(* IEC 61131-3 sources: rusty/tests/lit/single/arithmetic, 5 files *)

(* ---- addition.st ---- *)
// RUN: (%COMPILE %s && %RUN) | %CHECK %s
// CHECK: 10
FUNCTION main
    VAR
        x : DINT;
        y : DINT;
    END_VAR

    x := 5;
    y := 5;
    printf('%d$N', x + y);
END_FUNCTION

(* ---- integer_overflow.st ---- *)
// RUN: (%COMPILE %s && %RUN) | %CHECK %s
FUNCTION main
    VAR
        var_sint    : SINT;
        var_int     : INT;
        var_dint    : DINT;
        var_lint    : LINT;

        var_usint   : USINT;
        var_uint    : UINT;
        var_udint   : UDINT;
        var_ulint   : ULINT;
    END_VAR

    // Set max values
    // 8-bit [(2^7)-1]/[(2^8)-1]
    var_sint := 127;                    // Min: -128
    var_usint := 255;                   // Min: 0

    // 16-bit [(2^15)-1]/[(2^16)-1]
    var_int := 32767;                   // Min: -32768
    var_uint := 65535;                  // Min: 0

    // 32-bit [(2^31)-1]/[(2^31)-1]
    var_dint := 2147483647;             // Min: -2147483648
    var_udint := 4294967295;            // Min: 0

    // 64-bit [(2^63)-1]/[(2^64)-1]
    var_lint := 9223372036854775807;    // Min: -9223372036854775808
    var_ulint := 18446744073709551615;  // Min: 0

    // Print and check values
    printf('%d$N', var_sint);       // CHECK: 127
    printf('%d$N', var_int);        // CHECK-NEXT: 32767
    printf('%d$N', var_dint);       // CHECK-NEXT: 2147483647
    printf('%lld$N', var_lint);     // CHECK-NEXT: 9223372036854775807

    printf('%u$N', var_usint);      // CHECK-NEXT: 255
    printf('%u$N', var_uint);       // CHECK-NEXT: 65535
    printf('%u$N', var_udint);      // CHECK-NEXT: 4294967295
    printf('%llu$N', var_ulint);    // CHECK-NEXT: 18446744073709551615

    // Print overflow values
    var_sint := var_sint + 1;
    var_int := var_int + 1;
    var_dint := var_dint + 1;
    var_lint := var_lint + 1;

    var_usint := var_usint + 1;
    var_uint := var_uint + 1;
    var_udint := var_udint + 1;
    var_ulint := var_ulint + 1;

    printf('%d$N', var_sint);       // CHECK: -128
    printf('%d$N', var_int);        // CHECK-NEXT: -32768
    printf('%d$N', var_dint);       // CHECK-NEXT: -2147483648
    printf('%lld$N', var_lint);     // CHECK-NEXT: -9223372036854775808

    printf('%u$N', var_usint);      // CHECK-NEXT: 0
    printf('%u$N', var_uint);       // CHECK-NEXT: 0
    printf('%u$N', var_udint);      // CHECK-NEXT: 0
    printf('%llu$N', var_ulint);    // CHECK-NEXT: 0

END_FUNCTION

(* ---- integer_overflow_with_real_cast.st ---- *)
// RUN: (%COMPILE %s && %RUN) | %CHECK %s
FUNCTION main
    VAR
        var_int     : INT;
    END_VAR

    printf('%d$N', var_int); // CHECK: 0

    // Cast the REAL value to INT
    var_int := REAL_TO_INT(70_000.4);

    printf('%d$N', var_int); // CHECK: 32767

END_FUNCTION

(* ---- sqrt.st ---- *)
// RUN: (%COMPILE %s && %RUN) | %CHECK %s
// CHECK: 2
FUNCTION main
    VAR
        res : LREAL;
    END_VAR
    printf('%d$N', REAL_TO_DINT(SQRT(4.0)));
END_FUNCTION

(* ---- unsigned_with_literal.st ---- *)
// RUN: (%COMPILE %s && %RUN) | %CHECK %s

// An integer literal takes the type of an unsigned operand of 32 or 64 bits, so the operation stays unsigned
FUNCTION main : DINT
    VAR
        udintValue : UDINT := 4000000000;
        dwordValue : DWORD := 16#FFFFFFFF;
        ulintValue : ULINT := 18446744073709551615;
        ulintResult : ULINT;
        usintValue : USINT := 0;
        dintValue : DINT := -7;
    END_VAR

    // CHECK: 2000000000
    printf('%u$N', udintValue / 2);
    // CHECK: 3
    printf('%u$N', udintValue MOD 7);
    // CHECK: 1
    printf('%u$N', 4000000001 MOD udintValue);
    // CHECK: 2147483647
    printf('%u$N', dwordValue / 2);
    // CHECK: 0
    printf('%u$N', dwordValue MOD 3);
    // CHECK: 9223372036854775807
    printf('%llu$N', ulintValue / 2);

    ulintResult := udintValue + 1;
    // CHECK: 4000000001
    printf('%llu$N', ulintResult);

    // Smaller unsigned and signed operands are not affected
    // CHECK: -1
    printf('%d$N', usintValue - 1);
    // CHECK: -3
    printf('%d$N', dintValue / 2);
END_FUNCTION
